// TIA Portal V20 export
// export: Created 2026-10-12T05:42:32.6403764Z, ExportSetting WithDefaults, DisplayName Totally Integrated Automation Portal, DisplayVersion V20, DisplayName TIA Portal Openness, DisplayVersion V20, DisplayName TIA Portal Teamcenter Gateway, DisplayVersion V20, DisplayName TIA Portal Version Control Interface, DisplayVersion V20, DisplayName SINAMICS Startdrive Advanced, DisplayVersion V20 SP1 Update 2, DisplayName SINAMICS Startdrive G110M, G120, G120C, G120D, G120P, G115D, DisplayVersion V20 SP1 Update 2, DisplayName SINAMICS Startdrive G130, G150, S120, S150, SINAMICS MV, G220, S200, S210, DisplayVersion V20 SP1 Update 2, DisplayName STEP 7 Professional, DisplayVersion V20, DisplayName STEP 7 Safety, DisplayVersion V20, DisplayName WinCC Basic/Comfort/Advanced, DisplayVersion V20, DisplayName WinCC Professional, DisplayVersion V20, DisplayName WinCC Unified, DisplayVersion V20
FUNCTION "FRK_SeqStep" : Void   // FC129, SCL
{ S7_Optimized_Access := 'TRUE' }
VERSION : 0.1
// stored: AutoNumber true, IsIECCheckEnabled false, SetENOAutomatically false, UDAEnableTagReadback false
   VAR_INPUT
      StepNo : DInt;
      StepName : String;
   END_VAR
   VAR_IN_OUT
      Seq : "FRK_SequenceCtx";
      Row : "FRK_SequenceRow";
   END_VAR
BEGIN

   IF #Seq.RecordedStep <> #StepNo THEN
       #Seq.Visit := #Seq.Visit + 1;
       #Seq.Elapsed := T#0ms;
       #Seq.DelayElapsed := T#0ms;
       #Seq.RecordedStep := #StepNo;
       #Seq.Warned := FALSE;
   END_IF;
   #Seq.Step := #StepNo;
   #Seq.StepName := #StepName;
   #Row.StepNo := #StepNo;
   #Row.Visited := TRUE;
   #Row.LastDuration := #Seq.Elapsed;
END_FUNCTION
